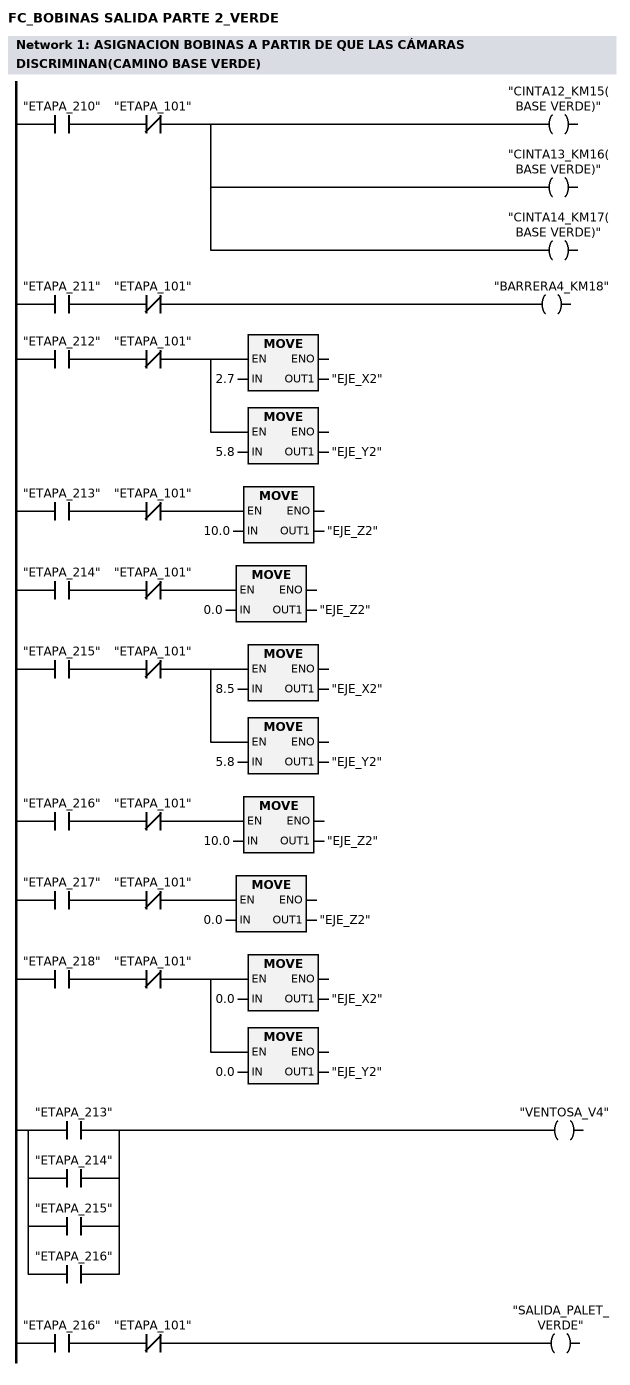
   RUNG wire#powerrail
      Contact( "ETAPA_210" )
      I_Contact( "ETAPA_101" )
      wire#w1
      Coil( "CINTA12_KM15(BASE VERDE)" )
   END_RUNG
   RUNG wire#w1
      Coil( "CINTA13_KM16(BASE VERDE)" )
   END_RUNG
   RUNG wire#w1
      Coil( "CINTA14_KM17(BASE VERDE)" )
   END_RUNG
   RUNG wire#powerrail
      Contact( "ETAPA_211" )
      I_Contact( "ETAPA_101" )
      Coil( "BARRERA4_KM18" )
   END_RUNG
   RUNG wire#powerrail
      Contact( "ETAPA_212" )
      I_Contact( "ETAPA_101" )
      wire#w2
      Move(in := 2.7, out1 => "EJE_X2")
   END_RUNG
   RUNG wire#w2
      Move(in := 5.8, out1 => "EJE_Y2")
   END_RUNG
   RUNG wire#powerrail
      Contact( "ETAPA_213" )
      I_Contact( "ETAPA_101" )
      Move(in := 10.0, out1 => "EJE_Z2")
   END_RUNG
   RUNG wire#powerrail
      Contact( "ETAPA_214" )
      I_Contact( "ETAPA_101" )
      Move(in := 0.0, out1 => "EJE_Z2")
   END_RUNG
   RUNG wire#powerrail
      Contact( "ETAPA_215" )
      I_Contact( "ETAPA_101" )
      wire#w3
      Move(in := 8.5, out1 => "EJE_X2")
   END_RUNG
   RUNG wire#w3
      Move(in := 5.8, out1 => "EJE_Y2")
   END_RUNG
   RUNG wire#powerrail
      Contact( "ETAPA_216" )
      I_Contact( "ETAPA_101" )
      Move(in := 10.0, out1 => "EJE_Z2")
   END_RUNG
   RUNG wire#powerrail
      Contact( "ETAPA_217" )
      I_Contact( "ETAPA_101" )
      Move(in := 0.0, out1 => "EJE_Z2")
   END_RUNG
   RUNG wire#powerrail
      Contact( "ETAPA_218" )
      I_Contact( "ETAPA_101" )
      wire#w4
      Move(in := 0.0, out1 => "EJE_X2")
   END_RUNG
   RUNG wire#w4
      Move(in := 0.0, out1 => "EJE_Y2")
   END_RUNG
   RUNG wire#powerrail
      Contact( "ETAPA_213" )
      wire#w5
      Coil( "VENTOSA_V4" )
   END_RUNG
   RUNG wire#powerrail
      Contact( "ETAPA_214" )
   END_RUNG wire#w5
   RUNG wire#powerrail
      Contact( "ETAPA_215" )
   END_RUNG wire#w5
   RUNG wire#powerrail
      Contact( "ETAPA_216" )
   END_RUNG wire#w5
   RUNG wire#powerrail
      Contact( "ETAPA_216" )
      I_Contact( "ETAPA_101" )
      Coil( "SALIDA_PALET_VERDE" )
   END_RUNG
   // the same network as SCL:
   "CINTA12_KM15(BASE VERDE)" := "ETAPA_210" AND NOT "ETAPA_101";
   "CINTA13_KM16(BASE VERDE)" := "CINTA12_KM15(BASE VERDE)";
   "CINTA14_KM17(BASE VERDE)" := "CINTA12_KM15(BASE VERDE)";
   "BARRERA4_KM18" := "ETAPA_211" AND NOT "ETAPA_101";
   IF "ETAPA_212" AND NOT "ETAPA_101" THEN
       "EJE_X2" := 2.7;
       "EJE_Y2" := 5.8;
   END_IF;
   IF "ETAPA_213" AND NOT "ETAPA_101" THEN "EJE_Z2" := 10.0; END_IF;
   IF "ETAPA_214" AND NOT "ETAPA_101" THEN "EJE_Z2" := 0.0; END_IF;
   IF "ETAPA_215" AND NOT "ETAPA_101" THEN
       "EJE_X2" := 8.5;
       "EJE_Y2" := 5.8;
   END_IF;
   IF "ETAPA_216" AND NOT "ETAPA_101" THEN "EJE_Z2" := 10.0; END_IF;
   IF "ETAPA_217" AND NOT "ETAPA_101" THEN "EJE_Z2" := 0.0; END_IF;
   IF "ETAPA_218" AND NOT "ETAPA_101" THEN
       "EJE_X2" := 0.0;
       "EJE_Y2" := 0.0;
   END_IF;
   "VENTOSA_V4" := "ETAPA_213" OR "ETAPA_214" OR "ETAPA_215" OR "ETAPA_216";
   "SALIDA_PALET_VERDE" := "ETAPA_216" AND NOT "ETAPA_101";
END_REGION
END_FUNCTION

FUNCTION "FC_SECUENCIA SALIDA PARTE 3_AZUL" : Void   // FC12, LAD
{ S7_Optimized_Access := 'TRUE' }
VERSION : 0.1
// N ESTE BLOQUE SE ENCUENTRA LA PROGRAMACIÓN DE LA SECUENCIA DESDE QUE LA PIEZA AZUL ES DEJADA EN EL PALET HASTA EL FINAL DEL PROCESO ALMACENANDOLA EN EL ALMACÉN
   VAR_TEMP   // added for the SCL form of the ladder/FBD networks
      _w1 : Bool;
   END_VAR
BEGIN

REGION Network 1: SECUENCIA DEL PROCESO DE SALIDA PARTE 3 (CAMINO BASE AZUL)
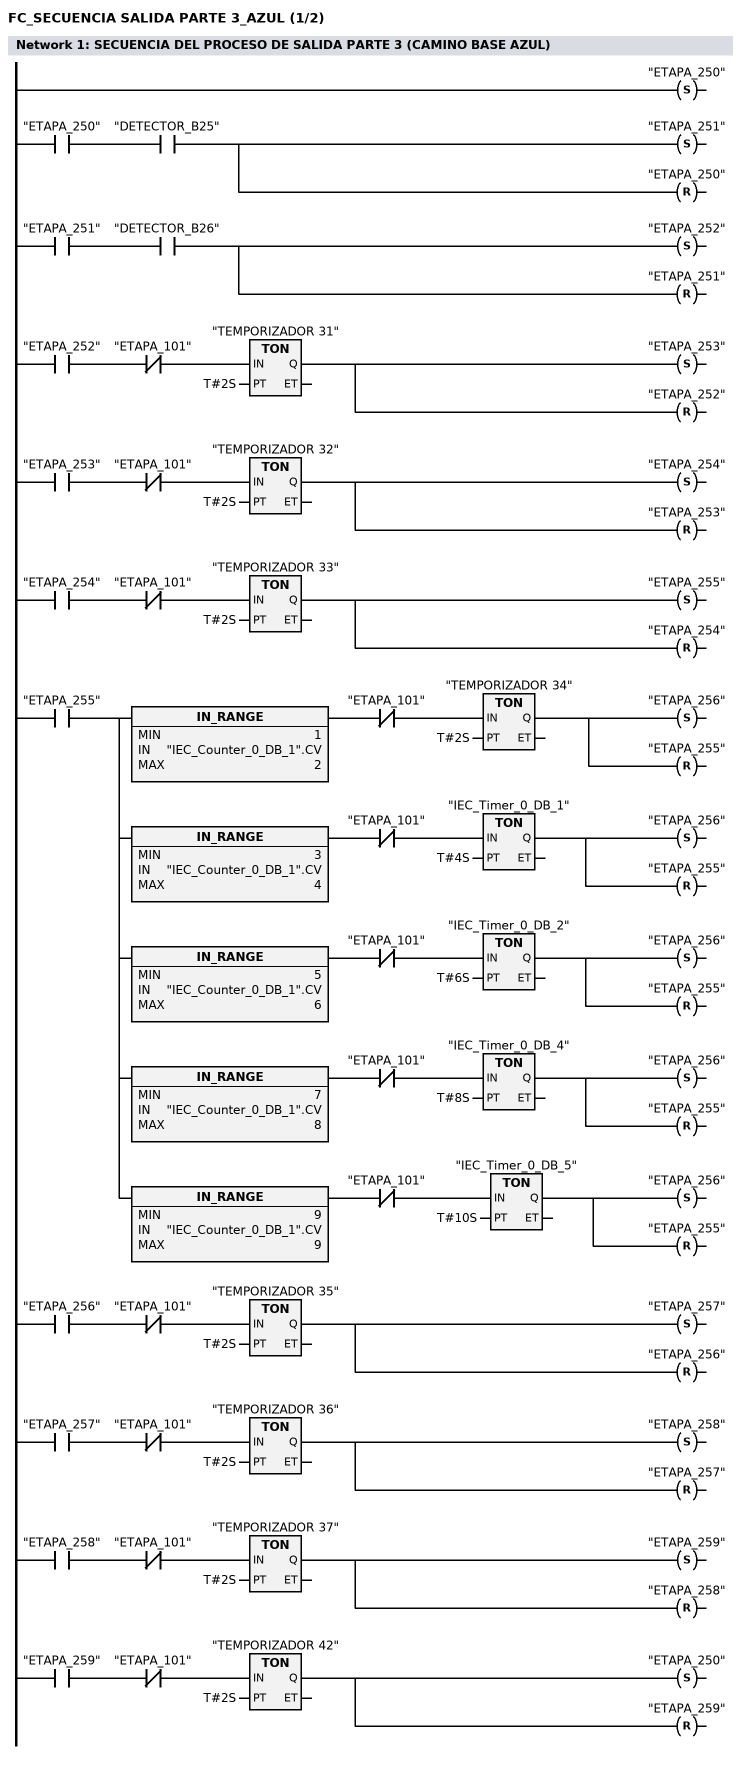
   "ETAPA_250" := TRUE;
   IF "ETAPA_250" AND "DETECTOR_B25" THEN
       "ETAPA_251" := TRUE;
       "ETAPA_250" := FALSE;
   END_IF;
   IF "ETAPA_251" AND "DETECTOR_B26" THEN
       "ETAPA_252" := TRUE;
       "ETAPA_251" := FALSE;
   END_IF;
   "TEMPORIZADOR 31".TON(IN := "ETAPA_252" AND NOT "ETAPA_101", PT := T#2S);
   IF "TEMPORIZADOR 31".Q THEN
       "ETAPA_253" := TRUE;
       "ETAPA_252" := FALSE;
   END_IF;
   "TEMPORIZADOR 32".TON(IN := "ETAPA_253" AND NOT "ETAPA_101", PT := T#2S);
   IF "TEMPORIZADOR 32".Q THEN
       "ETAPA_254" := TRUE;
       "ETAPA_253" := FALSE;
   END_IF;
   "TEMPORIZADOR 33".TON(IN := "ETAPA_254" AND NOT "ETAPA_101", PT := T#2S);
   IF "TEMPORIZADOR 33".Q THEN
       "ETAPA_255" := TRUE;
       "ETAPA_254" := FALSE;
   END_IF;
   "TEMPORIZADOR 34".TON(IN := "ETAPA_255" AND (1 <= "IEC_Counter_0_DB_1".CV) AND ("IEC_Counter_0_DB_1".CV <= 2) AND NOT "ETAPA_101",
                         PT := T#2S);
   IF "TEMPORIZADOR 34".Q THEN "ETAPA_256" := TRUE; END_IF;
   #_w1 := "ETAPA_255";
   IF "TEMPORIZADOR 34".Q THEN "ETAPA_255" := FALSE; END_IF;
   "IEC_Timer_0_DB_1".TON(IN := #_w1 AND (3 <= "IEC_Counter_0_DB_1".CV) AND ("IEC_Counter_0_DB_1".CV <= 4) AND NOT "ETAPA_101",
                          PT := T#4S);
   IF "IEC_Timer_0_DB_1".Q THEN
       "ETAPA_256" := TRUE;
       "ETAPA_255" := FALSE;
   END_IF;
   "IEC_Timer_0_DB_2".TON(IN := #_w1 AND (5 <= "IEC_Counter_0_DB_1".CV) AND ("IEC_Counter_0_DB_1".CV <= 6) AND NOT "ETAPA_101",
                          PT := T#6S);
   IF "IEC_Timer_0_DB_2".Q THEN
       "ETAPA_256" := TRUE;
       "ETAPA_255" := FALSE;
   END_IF;
   "IEC_Timer_0_DB_4".TON(IN := #_w1 AND (7 <= "IEC_Counter_0_DB_1".CV) AND ("IEC_Counter_0_DB_1".CV <= 8) AND NOT "ETAPA_101",
                          PT := T#8S);
   IF "IEC_Timer_0_DB_4".Q THEN
       "ETAPA_256" := TRUE;
       "ETAPA_255" := FALSE;
   END_IF;
   "IEC_Timer_0_DB_5".TON(IN := #_w1 AND (9 <= "IEC_Counter_0_DB_1".CV) AND ("IEC_Counter_0_DB_1".CV <= 9) AND NOT "ETAPA_101",
                          PT := T#10S);
   IF "IEC_Timer_0_DB_5".Q THEN
       "ETAPA_256" := TRUE;
       "ETAPA_255" := FALSE;
   END_IF;
   "TEMPORIZADOR 35".TON(IN := "ETAPA_256" AND NOT "ETAPA_101", PT := T#2S);
   IF "TEMPORIZADOR 35".Q THEN
       "ETAPA_257" := TRUE;
       "ETAPA_256" := FALSE;
   END_IF;
   "TEMPORIZADOR 36".TON(IN := "ETAPA_257" AND NOT "ETAPA_101", PT := T#2S);
   IF "TEMPORIZADOR 36".Q THEN
       "ETAPA_258" := TRUE;
       "ETAPA_257" := FALSE;
   END_IF;
   "TEMPORIZADOR 37".TON(IN := "ETAPA_258" AND NOT "ETAPA_101", PT := T#2S);
   IF "TEMPORIZADOR 37".Q THEN
       "ETAPA_259" := TRUE;
       "ETAPA_258" := FALSE;
   END_IF;
   "TEMPORIZADOR 42".TON(IN := "ETAPA_259" AND NOT "ETAPA_101", PT := T#2S);
   IF "TEMPORIZADOR 42".Q THEN
       "ETAPA_250" := TRUE;
       "ETAPA_259" := FALSE;
   END_IF;
END_REGION

REGION Network 2: PROGRAMACIÓN VISUALIZACIÓN ALMACENAMIENTO EN HMI
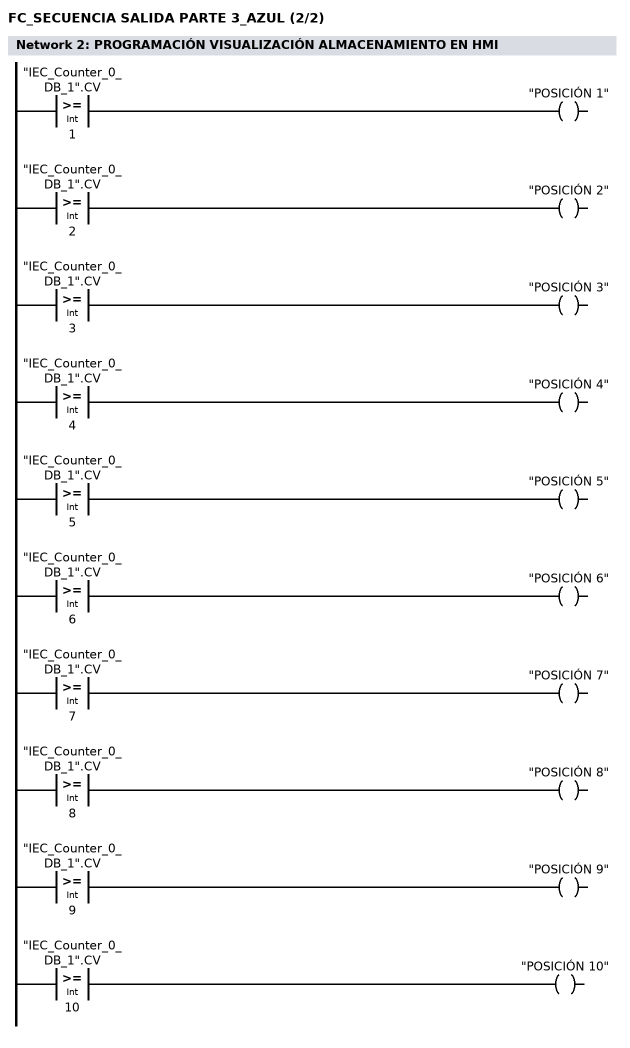
   RUNG wire#powerrail
      { S7_Templates := "SrcType := Int" } GE_Contact(in1 := "IEC_Counter_0_DB_1".CV, in2 := 1)
      Coil( "POSICIÓN 1" )
   END_RUNG
   RUNG wire#powerrail
      { S7_Templates := "SrcType := Int" } GE_Contact(in1 := "IEC_Counter_0_DB_1".CV, in2 := 2)
      Coil( "POSICIÓN 2" )
   END_RUNG
   RUNG wire#powerrail
      { S7_Templates := "SrcType := Int" } GE_Contact(in1 := "IEC_Counter_0_DB_1".CV, in2 := 3)
      Coil( "POSICIÓN 3" )
   END_RUNG
   RUNG wire#powerrail
      { S7_Templates := "SrcType := Int" } GE_Contact(in1 := "IEC_Counter_0_DB_1".CV, in2 := 4)
      Coil( "POSICIÓN 4" )
   END_RUNG
   RUNG wire#powerrail
      { S7_Templates := "SrcType := Int" } GE_Contact(in1 := "IEC_Counter_0_DB_1".CV, in2 := 5)
      Coil( "POSICIÓN 5" )
   END_RUNG
   RUNG wire#powerrail
      { S7_Templates := "SrcType := Int" } GE_Contact(in1 := "IEC_Counter_0_DB_1".CV, in2 := 6)
      Coil( "POSICIÓN 6" )
   END_RUNG
   RUNG wire#powerrail
      { S7_Templates := "SrcType := Int" } GE_Contact(in1 := "IEC_Counter_0_DB_1".CV, in2 := 7)
      Coil( "POSICIÓN 7" )
   END_RUNG
   RUNG wire#powerrail
      { S7_Templates := "SrcType := Int" } GE_Contact(in1 := "IEC_Counter_0_DB_1".CV, in2 := 8)
      Coil( "POSICIÓN 8" )
   END_RUNG
   RUNG wire#powerrail
      { S7_Templates := "SrcType := Int" } GE_Contact(in1 := "IEC_Counter_0_DB_1".CV, in2 := 9)
      Coil( "POSICIÓN 9" )
   END_RUNG
   RUNG wire#powerrail
      { S7_Templates := "SrcType := Int" } GE_Contact(in1 := "IEC_Counter_0_DB_1".CV, in2 := 10)
      Coil( "POSICIÓN 10" )
   END_RUNG
   // the same network as SCL:
   "POSICIÓN 1" := "IEC_Counter_0_DB_1".CV >= 1;
   "POSICIÓN 2" := "IEC_Counter_0_DB_1".CV >= 2;
   "POSICIÓN 3" := "IEC_Counter_0_DB_1".CV >= 3;
   "POSICIÓN 4" := "IEC_Counter_0_DB_1".CV >= 4;
   "POSICIÓN 5" := "IEC_Counter_0_DB_1".CV >= 5;
   "POSICIÓN 6" := "IEC_Counter_0_DB_1".CV >= 6;
   "POSICIÓN 7" := "IEC_Counter_0_DB_1".CV >= 7;
   "POSICIÓN 8" := "IEC_Counter_0_DB_1".CV >= 8;
   "POSICIÓN 9" := "IEC_Counter_0_DB_1".CV >= 9;
   "POSICIÓN 10" := "IEC_Counter_0_DB_1".CV >= 10;
END_REGION
END_FUNCTION

FUNCTION "FC_BOBINAS SALIDA PARTE 3_AZUL" : Void   // FC13, LAD
{ S7_Optimized_Access := 'TRUE' }
VERSION : 0.1
// EN ESTE BLOQUE SE ENCUENTRA LA ASIGNACIÓN DE CADA ETAPA CON EL ACTUADOR QUE CORRESPONDE, DESDE QUE LAS PIEZAS AZULES SON DEJADAS EN EL PALET HASTA QUE ACABA EL PROCESO DEJANDOLAS EN EL ALMCACEN
   VAR_TEMP   // added for the SCL form of the ladder/FBD networks
      _w1 : Bool;
   END_VAR
BEGIN

REGION Network 1: ASIGNACION BOBINAS A PARTIR DE QUE SON DEJADAS EN EL PALET(CAMINO BASE AZUL)
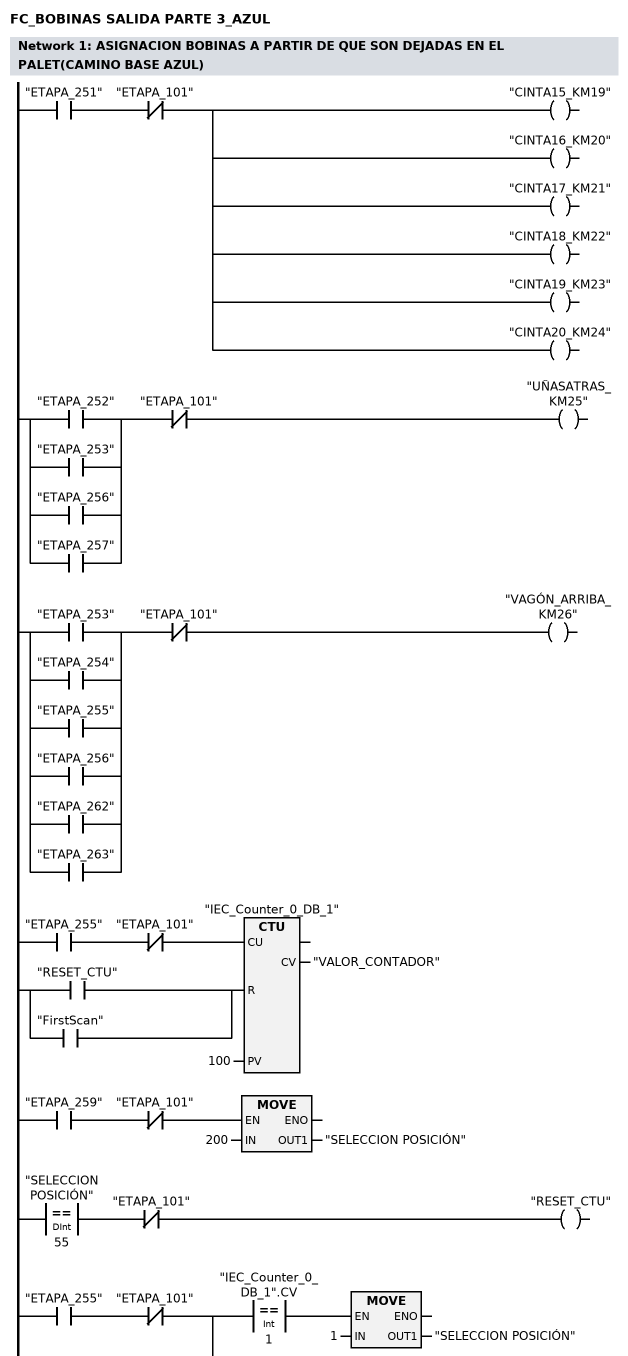
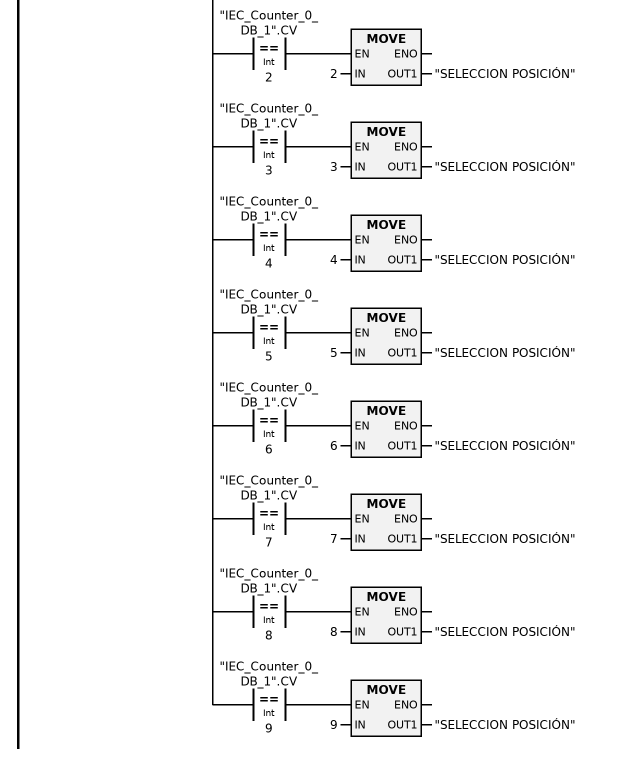
   "CINTA15_KM19" := "ETAPA_251" AND NOT "ETAPA_101";
   "CINTA16_KM20" := "CINTA15_KM19";
   "CINTA17_KM21" := "CINTA15_KM19";
   "CINTA18_KM22" := "CINTA15_KM19";
   "CINTA19_KM23" := "CINTA15_KM19";
   "CINTA20_KM24" := "CINTA15_KM19";
   "UÑASATRAS_KM25" := ("ETAPA_252" OR "ETAPA_253" OR "ETAPA_256" OR "ETAPA_257") AND NOT "ETAPA_101";
   "VAGÓN_ARRIBA_KM26" := ("ETAPA_253" OR "ETAPA_254" OR "ETAPA_255" OR "ETAPA_256" OR "ETAPA_262" OR "ETAPA_263") AND NOT "ETAPA_101";
   "IEC_Counter_0_DB_1".CTU(CU := "ETAPA_255" AND NOT "ETAPA_101",
                           R := "RESET_CTU" OR "FirstScan",
                           PV := 100,
                           CV => "VALOR_CONTADOR");
   IF "ETAPA_259" AND NOT "ETAPA_101" THEN "SELECCION POSICIÓN" := 200; END_IF;
   "RESET_CTU" := ("SELECCION POSICIÓN" = 55) AND NOT "ETAPA_101";
   #_w1 := "ETAPA_255" AND NOT "ETAPA_101";
   IF #_w1 AND ("IEC_Counter_0_DB_1".CV = 1) THEN "SELECCION POSICIÓN" := 1; END_IF;
   IF #_w1 AND ("IEC_Counter_0_DB_1".CV = 2) THEN "SELECCION POSICIÓN" := 2; END_IF;
   IF #_w1 AND ("IEC_Counter_0_DB_1".CV = 3) THEN "SELECCION POSICIÓN" := 3; END_IF;
   IF #_w1 AND ("IEC_Counter_0_DB_1".CV = 4) THEN "SELECCION POSICIÓN" := 4; END_IF;
   IF #_w1 AND ("IEC_Counter_0_DB_1".CV = 5) THEN "SELECCION POSICIÓN" := 5; END_IF;
   IF #_w1 AND ("IEC_Counter_0_DB_1".CV = 6) THEN "SELECCION POSICIÓN" := 6; END_IF;
   IF #_w1 AND ("IEC_Counter_0_DB_1".CV = 7) THEN "SELECCION POSICIÓN" := 7; END_IF;
   IF #_w1 AND ("IEC_Counter_0_DB_1".CV = 8) THEN "SELECCION POSICIÓN" := 8; END_IF;
   IF #_w1 AND ("IEC_Counter_0_DB_1".CV = 9) THEN "SELECCION POSICIÓN" := 9; END_IF;
END_REGION
END_FUNCTION

FUNCTION "FC_SECUENCIA SALIDA PARTE 3_VERDE" : Void   // FC14, LAD
{ S7_Optimized_Access := 'TRUE' }
VERSION : 0.1
// N ESTE BLOQUE SE ENCUENTRA LA PROGRAMACIÓN DE LA SECUENCIA DESDE QUE LA PIEZA VERDE ES DEJADA EN EL PALET HASTA EL FINAL DEL PROCESO ALMACENANDOLA EN EL ALMACÉN
BEGIN

REGION Network 1: SECUENCIA DEL PROCESO DE SALIDA PARTE 3 (CAMINO BASE VERDE)
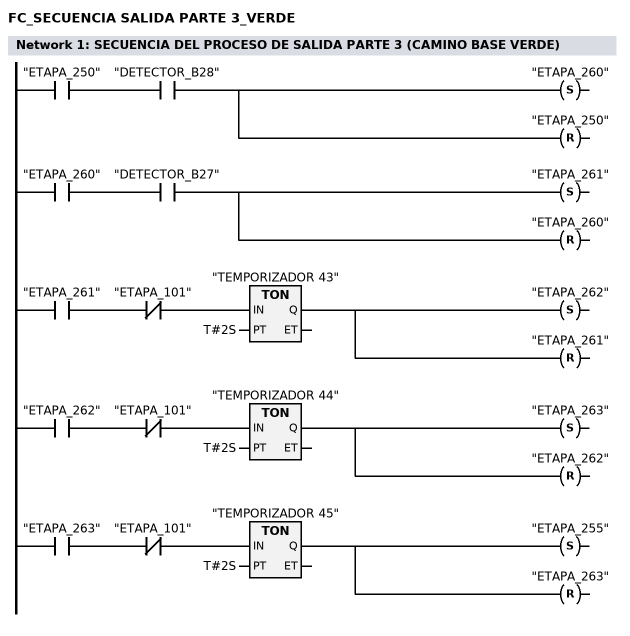
   IF "ETAPA_250" AND "DETECTOR_B28" THEN
       "ETAPA_260" := TRUE;
       "ETAPA_250" := FALSE;
   END_IF;
   IF "ETAPA_260" AND "DETECTOR_B27" THEN
       "ETAPA_261" := TRUE;
       "ETAPA_260" := FALSE;
   END_IF;
   "TEMPORIZADOR 43".TON(IN := "ETAPA_261" AND NOT "ETAPA_101", PT := T#2S);
   IF "TEMPORIZADOR 43".Q THEN
       "ETAPA_262" := TRUE;
       "ETAPA_261" := FALSE;
   END_IF;
   "TEMPORIZADOR 44".TON(IN := "ETAPA_262" AND NOT "ETAPA_101", PT := T#2S);
   IF "TEMPORIZADOR 44".Q THEN
       "ETAPA_263" := TRUE;
       "ETAPA_262" := FALSE;
   END_IF;
   "TEMPORIZADOR 45".TON(IN := "ETAPA_263" AND NOT "ETAPA_101", PT := T#2S);
   IF "TEMPORIZADOR 45".Q THEN
       "ETAPA_255" := TRUE;
       "ETAPA_263" := FALSE;
   END_IF;
END_REGION
END_FUNCTION

FUNCTION "FC_BOBINAS SALIDA PARTE 3_VERDE" : Void   // FC15, LAD
{ S7_Optimized_Access := 'TRUE' }
VERSION : 0.1
// EN ESTE BLOQUE SE ENCUENTRA LA ASIGNACIÓN DE CADA ETAPA CON EL ACTUADOR QUE CORRESPONDE, DESDE QUE LAS PIEZAS VERDES SON DEJADAS EN EL PALET HASTA QUE ACABA EL PROCESO DEJANDOLAS EN EL ALMCACEN
BEGIN

REGION Network 1: ASIGNACION BOBINAS A PARTIR DE QUE SON DEJADAS EN EL PALET(CAMINO BASE AZUL)
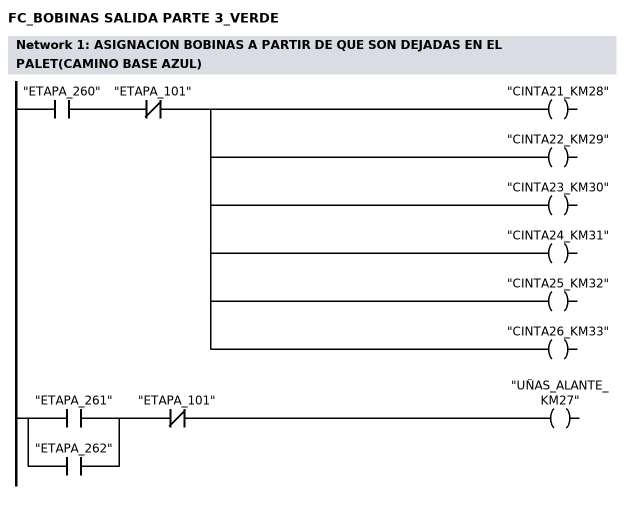
   RUNG wire#powerrail
      Contact( "ETAPA_260" )
      I_Contact( "ETAPA_101" )
      wire#w1
      Coil( "CINTA21_KM28" )
   END_RUNG
   RUNG wire#w1
      Coil( "CINTA22_KM29" )
   END_RUNG
   RUNG wire#w1
      Coil( "CINTA23_KM30" )
   END_RUNG
   RUNG wire#w1
      Coil( "CINTA24_KM31" )
   END_RUNG
   RUNG wire#w1
      Coil( "CINTA25_KM32" )
   END_RUNG
   RUNG wire#w1
      Coil( "CINTA26_KM33" )
   END_RUNG
   RUNG wire#powerrail
      Contact( "ETAPA_261" )
      wire#w2
      I_Contact( "ETAPA_101" )
      Coil( "UÑAS_ALANTE_KM27" )
   END_RUNG
   RUNG wire#powerrail
      Contact( "ETAPA_262" )
   END_RUNG wire#w2
   // the same network as SCL:
   "CINTA21_KM28" := "ETAPA_260" AND NOT "ETAPA_101";
   "CINTA22_KM29" := "CINTA21_KM28";
   "CINTA23_KM30" := "CINTA21_KM28";
   "CINTA24_KM31" := "CINTA21_KM28";
   "CINTA25_KM32" := "CINTA21_KM28";
   "CINTA26_KM33" := "CINTA21_KM28";
   "UÑAS_ALANTE_KM27" := ("ETAPA_261" OR "ETAPA_262") AND NOT "ETAPA_101";
END_REGION
END_FUNCTION

FUNCTION "MHJ-PLC-Lab-Function-S71200" : Void   // FC9000, SCL
{ S7_Optimized_Access := 'TRUE' }
VERSION : 0.1
   VAR_TEMP
      rdTimeReturn : Int;
      outputTime : DTL;
      SyncVal : Byte;
      forVal : Int;
      forVal_2 : Int;
      Value : Byte;
   END_VAR
   VAR CONSTANT
      CompVal : Byte := 16#34;
      Value_01 : Byte := 16#11;
      Value_01_DW : DWord := 16#A165_D992;
      Value_02_DW : DWord := 16#58BE_4401;
   END_VAR
BEGIN

   #Value:=PEEK(area := 16#82,
        dbNumber := 0,
        byteOffset := 511);
   #Value := #Value + 1;

   POKE(area := 16#82,
        dbNumber := 0,
        byteOffset := 511,
        value := #Value);

   POKE(area:=16#81,
        dbNumber:=0,
        byteOffset:=1016,
        value:=#Value_01_DW);
   POKE(area := 16#81,
        dbNumber := 0,
        byteOffset := 1020,
        value := #Value_02_DW);

   POKE(area := 16#81,
        dbNumber := 0,
        byteOffset := 511,
        value := B#16#00);

   FOR #forVal := 0 TO 120 DO
       FOR #forVal_2:=0 TO 10 DO
           #rdTimeReturn:=RD_SYS_T(#outputTime);
           #rdTimeReturn := WR_SYS_T(#outputTime);
           #rdTimeReturn := RD_SYS_T(#outputTime);
           #rdTimeReturn := WR_SYS_T(#outputTime);
       END_FOR;
       #SyncVal:= PEEK(area := 16#81,
                      dbNumber := 0,
                      byteOffset := 511);
       IF #SyncVal = #CompVal THEN
          GOTO M_1;
       END_IF;
   END_FOR;
   RETURN;

   M_1:
   POKE(area := 16#81,
        dbNumber := 0,
        byteOffset := 511,
        value := B#16#0);
END_FUNCTION

ORGANIZATION_BLOCK "Main"   // OB1, LAD, ProgramCycle
TITLE = "Main Program Sweep (Cycle)"
{ S7_Optimized_Access := 'TRUE' }
VERSION : 0.1
// EN ESTE BLOQUE TENEMOS LAS LLAMADAS AL MAIN DE LOS FC'S DEL PROCESO
   VAR_INPUT
      Initial_Call : Bool;   // Initial call of this OB
      Remanence : Bool;   // =True, if remanent data are available
   END_VAR
BEGIN

REGION Network 1
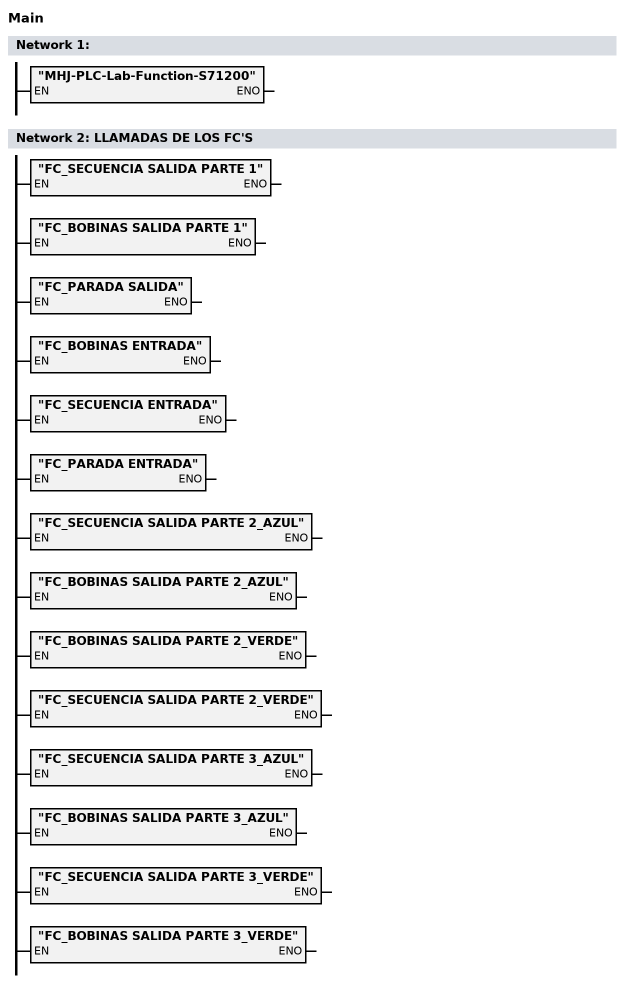
   RUNG wire#powerrail
      "MHJ-PLC-Lab-Function-S71200"()
   END_RUNG
   // the same network as SCL:
   "MHJ-PLC-Lab-Function-S71200"();
END_REGION

REGION Network 2: LLAMADAS DE LOS FC'S
   RUNG wire#powerrail
      "FC_SECUENCIA SALIDA PARTE 1"()
   END_RUNG
   RUNG wire#powerrail
      "FC_BOBINAS SALIDA PARTE 1"()
   END_RUNG
   RUNG wire#powerrail
      "FC_PARADA SALIDA"()
   END_RUNG
   RUNG wire#powerrail
      "FC_BOBINAS ENTRADA"()
   END_RUNG
   RUNG wire#powerrail
      "FC_SECUENCIA ENTRADA"()
   END_RUNG
   RUNG wire#powerrail
      "FC_PARADA ENTRADA"()
   END_RUNG
   RUNG wire#powerrail
      "FC_SECUENCIA SALIDA PARTE 2_AZUL"()
   END_RUNG
   RUNG wire#powerrail
      "FC_BOBINAS SALIDA PARTE 2_AZUL"()
   END_RUNG
   RUNG wire#powerrail
      "FC_BOBINAS SALIDA PARTE 2_VERDE"()
   END_RUNG
   RUNG wire#powerrail
      "FC_SECUENCIA SALIDA PARTE 2_VERDE"()
   END_RUNG
   RUNG wire#powerrail
      "FC_SECUENCIA SALIDA PARTE 3_AZUL"()
   END_RUNG
   RUNG wire#powerrail
      "FC_BOBINAS SALIDA PARTE 3_AZUL"()
   END_RUNG
   RUNG wire#powerrail
      "FC_SECUENCIA SALIDA PARTE 3_VERDE"()
   END_RUNG
   RUNG wire#powerrail
      "FC_BOBINAS SALIDA PARTE 3_VERDE"()
   END_RUNG
   // the same network as SCL:
   "FC_SECUENCIA SALIDA PARTE 1"();
   "FC_BOBINAS SALIDA PARTE 1"();
   "FC_PARADA SALIDA"();
   "FC_BOBINAS ENTRADA"();
   "FC_SECUENCIA ENTRADA"();
   "FC_PARADA ENTRADA"();
   "FC_SECUENCIA SALIDA PARTE 2_AZUL"();
   "FC_BOBINAS SALIDA PARTE 2_AZUL"();
   "FC_BOBINAS SALIDA PARTE 2_VERDE"();
   "FC_SECUENCIA SALIDA PARTE 2_VERDE"();
   "FC_SECUENCIA SALIDA PARTE 3_AZUL"();
   "FC_BOBINAS SALIDA PARTE 3_AZUL"();
   "FC_SECUENCIA SALIDA PARTE 3_VERDE"();
   "FC_BOBINAS SALIDA PARTE 3_VERDE"();
END_REGION
END_ORGANIZATION_BLOCK

ORGANIZATION_BLOCK "Startup"   // OB100, LAD, Startup
TITLE = "Complete Restart"
{ S7_Optimized_Access := 'TRUE' }
VERSION : 0.1
// EN ESTE BLOQUE SE ENCUENTRA EL RESET DE TODAS LAS ETAPAS
   VAR_INPUT
      LostRetentive : Bool;   // True if retentive data are lost
      LostRTC : Bool;   // True if date and time are lost
   END_VAR
BEGIN

REGION Network 1: RESET DE TODAS LAS ETAPAS
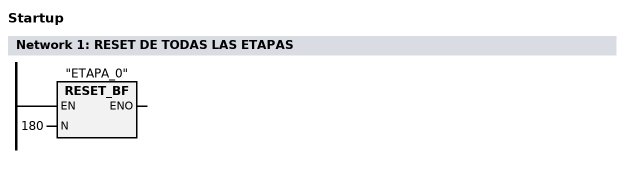
   // no SCL statement known for RBitfield: written as a call
   RESET_BF(operand := "ETAPA_0", n := 180);
END_REGION
END_ORGANIZATION_BLOCK

(* ===== HMI "HMI_RT_2" =====
system functions are stored by id; their names below are inferred from use
connection "HMI_Conexión_1": ETHERNET, S7_1200_OMS

HMI tags "Tabla de variables estándar"
   "POSICIÓN 1" : Bool = PLC "POSICIÓN 1" AT %M543.0, 1 s
   "POSICIÓN 2" : Bool = PLC "POSICIÓN 2" AT %M543.1, 1 s
   "POSICIÓN 3" : Bool = PLC "POSICIÓN 3" AT %M543.2, 1 s
   "POSICIÓN 4" : Bool = PLC "POSICIÓN 4" AT %M543.3, 1 s
   "POSICIÓN 5" : Bool = PLC "POSICIÓN 5" AT %M543.4, 1 s
   "POSICIÓN 6" : Bool = PLC "POSICIÓN 6" AT %M543.5, 1 s
   "POSICIÓN 7" : Bool = PLC "POSICIÓN 7" AT %M543.6, 1 s
   "POSICIÓN 8" : Bool = PLC "POSICIÓN 8" AT %M543.7, 1 s
   "POSICIÓN 9" : Bool = PLC "POSICIÓN 9" AT %M544.0, 1 s
   "POSICIÓN 10" : Bool = PLC "POSICIÓN 10" AT %M544.1, 1 s
   "VALOR_CONTADOR" : Int = PLC VALOR_CONTADOR AT %IW6, 1 s
   "VALOR_PROCESO_ENTRADA" : Int = PLC VALOR_PROCESO_ENTRADA AT %QW15, 1 s
   "MARCHA2_S5" : Bool = PLC MARCHA2_S5 AT %I2.5, 1 s
   "PARO2_S8" : Bool = PLC PARO2_S8 AT %I2.7, 1 s
   "RESET2_S14" : Bool = PLC RESET2_S14 AT %I4.2, 1 s
   "VALOR_PROCESO_SALIDA" : Int = PLC VALOR_PROCESO_SALIDA AT %QW20, 1 s
   "PULSADOR_S1" : Bool = PLC PULSADOR_S1 AT %I0.0, 1 s
   "PULSADOR_S2" : Bool = PLC PULSADOR_S2 AT %I0.1, 1 s
   "RESET1_S11" : Bool = PLC RESET1_S11 AT %I4.1, 1 s
   "MARCAA_VACIIA" : Bool = PLC MARCAA_VACIIA AT %M730.0, 1 s

text list "PROCESO ENTRADA": 1 'PROCESO EN MARCHA'; 2 'PROCESO PARADO'; 3 'PROCESO EN ALARMA'

text list "PROCESO SALIDA": 1 'PROCESO EN MARCHA'; 2 'PROCESO PARADO'; 3 'PROCESO EN ALARMA'

graphic list "VISUALIZACIÓN CAJA": 0 'Gráfico_17'; 1 'Gráfico_17'

graphic list "PROCESO ENTRADA GRAFICOS": 1 'Gráfico_18'; 2 'Gráfico_19'; 3 'Gráfico_20'

graphic list "PROCESO SALIDA GRAFICOS": 1 'Gráfico_18'; 2 'Gráfico_19'; 3 'Gráfico_20'

screen "INICIO" 1980x1080
   GraphicView "Visor de gráficos_2" at 13,80 size 119x103; Picture "Gráfico_13"
   DateTimeField "Campo de fecha y hora_1" at 0,0 size 234x62
   Button "Botón_1" at 7,73 size 145x105; TextOff 'Text'
      on Activate: ActivateScreen("INICIO", 0)
   Button "Botón_2" at 301,73 size 180x85; TextOff 'LOGIN'; PictureOff "vecteezy_rectangle-shape-buttons-in-green-colors-user-interface_14324191"
      on Click: function_a2a04561()
   Button "Botón_3" at 574,73 size 178x83; TextOn 'LONGOUT'; TextOff 'LONGOUT'; PictureOff "vecteezy_glossy-buttons-clipart-design-illustration_9342302"
      on Click: function_f23ef4c9()
   Button "Botón_4" at 863,80 size 228x83; TextOn 'PARAR RUNTIME'; TextOff 'PARAR RUNTIME'; PictureOff "vecteezy_glossy-buttons-clipart-design-illustration_9304864"
      on Click: StopRuntime(0)
   GraphicView "Visor de gráficos_3" at 1647,2 size 248x190; Picture "Gráfico_15"
   Button "Botón_5" at 344,945 size 289x85; TextOn 'CONTROL'; TextOff 'CONTROL'; PictureOff "vecteezy_rectangulo-de-sombra-rectangulo-neumorfico_11888129"; Authorization "CONTROL"
      on Press: function_efd93a16("CONTROL", 0, 191, -1, -1, 1)
   Button "Botón_6" at 1122,945 size 289x85; TextOn 'VISUALIZACIÓN'; TextOff 'VISUALIZACIÓN'; PictureOff "vecteezy_rectangulo-de-sombra-rectangulo-neumorfico_11888129"; Authorization "VISUALIZACIÓN"
      on Press: function_efd93a16("VISUALIZACIÓN", 0, 191, -1, -1, 1)
   GraphicView "Visor de gráficos_1" at 0,194 size 1979x751; Picture "Gráfico_21"

PopupScreen "CONTROL" 1980x752
   TextField "Campo de texto_1" at 781,26 size 532x77; Text 'CONTROL DEL PROCESO'
   Button "Botón_1" at 406,413 size 137x64; TextOff 'MARCHA'; PictureOff "vecteezy_glossy-buttons-clipart-design-illustration_9301007"
      on Press: function_b14e0dd5("MARCHA2_S5", 0)
   GraphicIOField "Campo ES gráfico_1" at 481,225 size 163x115; PictureList "PROCESO ENTRADA GRAFICOS"
      ProcessValue <- "VALOR_PROCESO_ENTRADA"
   SymbolicIOField "Campo ES simbólico_1" at 456,358 size 290x38; TextOff '0'; TextOn '1'; TextList "PROCESO ENTRADA"
      ProcessValue <- "VALOR_PROCESO_ENTRADA"
   Button "Botón_2" at 587,413 size 135x61; TextOn 'PARO'; TextOff 'PARO'; PictureOff "vecteezy_glossy-buttons-clipart-design-illustration_9342302"
      on Press: function_b14e0dd5("PARO2_S8", 0)
   Button "Botón_6" at 452,493 size 239x89; TextOn 'RESET'; TextOff 'RESET'; PictureOff "vecteezy_diseno-de-icono-de-forma_9266311"
      on Press: function_b14e0dd5("RESET2_S14", 0)
   TextField "Campo de texto_2" at 435,140 size 334x40; Text 'PROCESO DE ENTRADA'
   TextField "Campo de texto_3" at 1253,142 size 273x44; Text 'PROCESO DE SALIDA'
   GraphicIOField "Campo ES gráfico_2" at 1313,225 size 163x115; PictureList "PROCESO SALIDA GRAFICOS"
      ProcessValue <- "VALOR_PROCESO_SALIDA"
   Button "Botón_3" at 1239,413 size 137x64; TextOn 'MARCHA'; TextOff 'MARCHA'; PictureOff "vecteezy_glossy-buttons-clipart-design-illustration_9301007"
      on Press: function_b14e0dd5("PULSADOR_S1", 0)
   Button "Botón_4" at 1418,416 size 135x61; TextOn 'PARO'; TextOff 'PARO'; PictureOff "vecteezy_glossy-buttons-clipart-design-illustration_9342302"
      on Press: function_b14e0dd5("PULSADOR_S2", 0)
   Button "Botón_5" at 1280,493 size 239x89; TextOn 'RESET'; TextOff 'RESET'; PictureOff "vecteezy_diseno-de-icono-de-forma_9266311"
      on Press: function_b14e0dd5("RESET1_S11", 0)
   SymbolicIOField "Campo ES simbólico_2" at 1280,367 size 290x38; TextOn '1'; TextOff '0'; TextList "PROCESO SALIDA"
      ProcessValue <- "VALOR_PROCESO_ENTRADA"

PopupScreen "VISUALIZACIÓN" 1980x752
   Rectangle "Rectángulo_1" at 536,544 size 58x19
      Appearance <- "POSICIÓN 1"
   Rectangle "Rectángulo_2" at 615,544 size 58x19
      Appearance <- "POSICIÓN 2"
   Rectangle "Rectángulo_3" at 694,544 size 58x19
      Appearance <- "POSICIÓN 3"
   Rectangle "Rectángulo_4" at 773,544 size 58x19
      Appearance <- "POSICIÓN 4"
   Rectangle "Rectángulo_5" at 852,544 size 58x19
      Appearance <- "POSICIÓN 5"
   Rectangle "Rectángulo_6" at 931,544 size 58x19
      Appearance <- "POSICIÓN 6"
   Rectangle "Rectángulo_7" at 1010,544 size 58x19
      Appearance <- "POSICIÓN 7"
   Rectangle "Rectángulo_8" at 1089,544 size 58x19
      Appearance <- "POSICIÓN 8"
   Rectangle "Rectángulo_9" at 1168,544 size 58x19
      Appearance <- "POSICIÓN 9"
   Rectangle "Rectángulo_10" at 1247,544 size 58x19
      Appearance <- "POSICIÓN 10"
   GraphicView "Visor de gráficos_4" at 776,496 size 48x45; Picture "Gráfico_17"
      Visibility <- "POSICIÓN 4"
   GraphicView "Visor de gráficos_5" at 855,497 size 48x45; Picture "Gráfico_17"
      Visibility <- "POSICIÓN 5"
   GraphicView "Visor de gráficos_6" at 934,498 size 48x45; Picture "Gráfico_17"
      Visibility <- "POSICIÓN 6"
   GraphicView "Visor de gráficos_7" at 1013,499 size 48x45; Picture "Gráfico_17"
      Visibility <- "POSICIÓN 7"
   GraphicView "Visor de gráficos_8" at 1092,498 size 48x45; Picture "Gráfico_17"
      Visibility <- "POSICIÓN 8"
   GraphicView "Visor de gráficos_9" at 1171,499 size 48x45; Picture "Gráfico_17"
      Visibility <- "POSICIÓN 9"
   GraphicView "Visor de gráficos_10" at 1250,498 size 48x45; Picture "Gráfico_17"
      Visibility <- "POSICIÓN 10"
   GraphicView "Visor de gráficos_11" at 540,406 size 48x45; Picture "Gráfico_17"
      Visibility <- "MARCAA_VACIIA"
   GraphicView "Visor de gráficos_12" at 621,406 size 48x45; Picture "Gráfico_17"
      Visibility <- "MARCAA_VACIIA"
   GraphicView "Visor de gráficos_13" at 701,406 size 48x45; Picture "Gráfico_17"
      Visibility <- "MARCAA_VACIIA"
   GraphicView "Visor de gráficos_14" at 777,406 size 48x45; Picture "Gráfico_17"
      Visibility <- "MARCAA_VACIIA"
   GraphicView "Visor de gráficos_15" at 855,406 size 48x45; Picture "Gráfico_17"
      Visibility <- "MARCAA_VACIIA"
   GraphicView "Visor de gráficos_16" at 934,406 size 48x45; Picture "Gráfico_17"
      Visibility <- "MARCAA_VACIIA"
   GraphicView "Visor de gráficos_17" at 1012,406 size 48x45; Picture "Gráfico_17"
      Visibility <- "MARCAA_VACIIA"
   GraphicView "Visor de gráficos_18" at 1089,406 size 48x45; Picture "Gráfico_17"
      Visibility <- "MARCAA_VACIIA"
   GraphicView "Visor de gráficos_19" at 1168,406 size 48x45; Picture "Gráfico_17"
      Visibility <- "MARCAA_VACIIA"
   GraphicView "Visor de gráficos_20" at 1247,406 size 48x45; Picture "Gráfico_17"
      Visibility <- "MARCAA_VACIIA"
   GraphicView "Visor de gráficos_21" at 540,320 size 48x45; Picture "Gráfico_17"
      Visibility <- "MARCAA_VACIIA"
   GraphicView "Visor de gráficos_22" at 617,323 size 48x45; Picture "Gráfico_17"
      Visibility <- "MARCAA_VACIIA"
   GraphicView "Visor de gráficos_23" at 694,323 size 48x45; Picture "Gráfico_17"
      Visibility <- "MARCAA_VACIIA"
   GraphicView "Visor de gráficos_24" at 775,323 size 48x45; Picture "Gráfico_17"
      Visibility <- "MARCAA_VACIIA"
   GraphicView "Visor de gráficos_25" at 854,323 size 48x45; Picture "Gráfico_17"
      Visibility <- "MARCAA_VACIIA"
   GraphicView "Visor de gráficos_26" at 933,323 size 48x45; Picture "Gráfico_17"
      Visibility <- "MARCAA_VACIIA"
   GraphicView "Visor de gráficos_27" at 1012,323 size 48x45; Picture "Gráfico_17"
      Visibility <- "MARCAA_VACIIA"
   GraphicView "Visor de gráficos_28" at 1091,323 size 48x45; Picture "Gráfico_17"
      Visibility <- "MARCAA_VACIIA"
   GraphicView "Visor de gráficos_29" at 1170,323 size 48x45; Picture "Gráfico_17"
      Visibility <- "MARCAA_VACIIA"
   GraphicView "Visor de gráficos_30" at 1249,323 size 48x45; Picture "Gráfico_17"
      Visibility <- "MARCAA_VACIIA"
   GraphicView "Visor de gráficos_31" at 540,231 size 48x45; Picture "Gráfico_17"
      Visibility <- "MARCAA_VACIIA"
   GraphicView "Visor de gráficos_32" at 617,231 size 48x45; Picture "Gráfico_17"
      Visibility <- "MARCAA_VACIIA"
   GraphicView "Visor de gráficos_33" at 698,231 size 48x45; Picture "Gráfico_17"
      Visibility <- "MARCAA_VACIIA"
   GraphicView "Visor de gráficos_34" at 775,231 size 48x45; Picture "Gráfico_17"
      Visibility <- "MARCAA_VACIIA"
   GraphicView "Visor de gráficos_35" at 854,231 size 48x45; Picture "Gráfico_17"
      Visibility <- "MARCAA_VACIIA"
   GraphicView "Visor de gráficos_36" at 932,231 size 48x45; Picture "Gráfico_17"
      Visibility <- "MARCAA_VACIIA"
   GraphicView "Visor de gráficos_37" at 1013,231 size 48x45; Picture "Gráfico_17"
      Visibility <- "MARCAA_VACIIA"
   GraphicView "Visor de gráficos_38" at 1090,231 size 48x45; Picture "Gráfico_17"
      Visibility <- "MARCAA_VACIIA"
   GraphicView "Visor de gráficos_39" at 1171,230 size 48x45; Picture "Gráfico_17"
      Visibility <- "MARCAA_VACIIA"
   GraphicView "Visor de gráficos_40" at 1247,231 size 48x45; Picture "Gráfico_17"
      Visibility <- "MARCAA_VACIIA"
   GraphicView "Visor de gráficos_41" at 536,145 size 48x45; Picture "Gráfico_17"
      Visibility <- "MARCAA_VACIIA"
   GraphicView "Visor de gráficos_42" at 619,146 size 48x45; Picture "Gráfico_17"
      Visibility <- "MARCAA_VACIIA"
   GraphicView "Visor de gráficos_43" at 702,147 size 48x45; Picture "Gráfico_17"
      Visibility <- "MARCAA_VACIIA"
   GraphicView "Visor de gráficos_44" at 780,148 size 48x45; Picture "Gráfico_17"
      Visibility <- "MARCAA_VACIIA"
   GraphicView "Visor de gráficos_45" at 857,148 size 48x45; Picture "Gráfico_17"
      Visibility <- "MARCAA_VACIIA"
   GraphicView "Visor de gráficos_46" at 936,148 size 48x45; Picture "Gráfico_17"
      Visibility <- "MARCAA_VACIIA"
   GraphicView "Visor de gráficos_47" at 1016,148 size 48x45; Picture "Gráfico_17"
      Visibility <- "MARCAA_VACIIA"
   GraphicView "Visor de gráficos_48" at 1093,148 size 48x45; Picture "Gráfico_17"
      Visibility <- "MARCAA_VACIIA"
   GraphicView "Visor de gráficos_49" at 1171,148 size 48x45; Picture "Gráfico_17"
      Visibility <- "MARCAA_VACIIA"
   GraphicView "Visor de gráficos_50" at 1253,148 size 48x45; Picture "Gráfico_17"
      Visibility <- "MARCAA_VACIIA"
   TextField "Campo de texto_1" at 824,84 size 125x31; Text 'CONTADOR'
   IOField "Campo ES_1" at 957,84 size 96x32; FormatPattern 99
      ProcessValue <- "VALOR_CONTADOR"
   GraphicIOField "Campo ES gráfico_2" at 619,498 size 48x41; PictureList "VISUALIZACIÓN CAJA"
      ProcessValue <- "POSICIÓN 2"
      Visibility <- "POSICIÓN 2"
   GraphicIOField "Campo ES gráfico_3" at 698,499 size 48x41; PictureList "VISUALIZACIÓN CAJA"
      ProcessValue <- "POSICIÓN 3"
      Visibility <- "POSICIÓN 3"
   GraphicIOField "Campo ES gráfico_1" at 539,500 size 48x41; PictureList "VISUALIZACIÓN CAJA"
      ProcessValue <- "POSICIÓN 2"
      Visibility <- "POSICIÓN 1"
*)